(* IEC 61131-3 sources: structured-text/samples/unsupported/arrays, 10 files *)

(* ---- f.4.st ---- *)
FUNCTION_BLOCK STACK_INT
  VAR_INPUT PUSH, POP: BOOL;
            R1 : BOOL ;
            IN : INT ;
            N  : INT ;
  END_VAR
  VAR_OUTPUT EMPTY : BOOL := 1 ;
             OFLO  : BOOL := 0 ;
             OUT   : INT  := 0 ;
  END_VAR
  VAR STK : ARRAY[0..127] OF INT;
      NI : INT :=128  ;
      PTR : INT := -1 ;
  END_VAR

    IF R1 THEN
       OFLO := 0; EMPTY := 1; PTR := -1;
       NI := LIMIT (MN:=1,IN:=N,MX:=128); OUT := 0;
    ELSIF POP & NOT EMPTY THEN
       OFLO := 0; PTR := PTR-1; EMPTY := PTR < 0;
       IF EMPTY THEN OUT := 0;
       ELSE OUT := STK[PTR];
       END_IF ;
    ELSIF PUSH & NOT OFLO THEN
       EMPTY := 0; PTR := PTR+1; OFLO := (PTR = NI);
       IF NOT OFLO THEN OUT := IN ; STK[PTR] := IN;
       ELSE OUT := 0;
       END_IF ;
    END_IF ;
END_FUNCTION_BLOCK

(* ---- f.6.11.st ---- *)
FUNCTION_BLOCK DIFFEQ
   VAR_INPUT
     RUN : BOOL ;
     XIN : REAL ;
     A : ARRAY[1..127] OF REAL ;
     M : INT ;
     B : ARRAY[0..127] OF REAL ;
     N : INT ;
   END_VAR
   VAR_OUTPUT XOUT : REAL := 0.0 ; END_VAR
   VAR
     XI : ARRAY [0..127] OF REAL ;
     XO : ARRAY [0..127] OF REAL ;
     I : INT ;
   END_VAR
   XO[0] := XOUT ; XI[0] := XIN ;
   XOUT := B[0] * XIN ;
   IF RUN THEN
      FOR I := M TO 1 BY -1 DO
          XOUT := XOUT + A[I] * XO[I] ; XO[I] := XO[I-1];
      END_FOR;
      FOR I := N TO 1 BY -1 DO
          XOUT := XOUT + B[I] * XI[I] ; XI[I] := XI[I-1];
      END_FOR;
   ELSE
      FOR I := 1 TO M DO XO[I] := 0.0; END_FOR;
      FOR I := 1 TO N DO XI[I] := 0.0; END_FOR;
   END_IF ;
 END_FUNCTION_BLOCK

(* ---- f.6.2.st ---- *)
FUNCTION_BLOCK DELAY
  VAR_INPUT
    RUN : BOOL ;
    XIN : REAL ;
    N   : INT ;
  END_VAR
  VAR_OUTPUT XOUT : REAL; END_VAR
  VAR X : ARRAY [0..127]
               OF REAL;
      I, IXIN, IXOUT : INT := 0;
  END_VAR
  IF RUN THEN IXIN := MOD(IXIN + 1, 128) ; X[IXIN] := XIN ;
              IXOUT := MOD(IXOUT + 1, 128) ; XOUT := X[IXOUT];
  ELSE XOUT := XIN ; IXIN := N ; IXOUT := 0;
       FOR I := 0 TO N DO X[I] := XIN; END_FOR;
  END_IF ;
END_FUNCTION_BLOCK

(* ---- t17-4.st ---- *)
PROGRAM Test
	VAR
		INARY AT %IW6 ;
 		ARRAY [0..9] OF INT;
	END_VAR
END_PROGRAM

(* ---- t17-6.st ---- *)
PROGRAM Test
	VAR THREE :
		ARRAY[1..5,1..10,1..8] OF INT;
	END_VAR
END_PROGRAM

(* ---- t17-7.st ---- *)
PROGRAM Test
	VAR RETAIN RTBT:
  		ARRAY[1..2,1..3] OF INT;
	END_VAR
END_PROGRAM

(* ---- t18-4.st ---- *)
PROGRAM Test
	VAR OUTARY AT %QW6 :
 		ARRAY[0..9] OF INT := [10(1)];
	END_VAR
END_PROGRAM

(* ---- t18-6.st ---- *)
PROGRAM Test
	VAR
		BITS : ARRAY[0..7]
			OF BOOL := [1,1,0,0,0,1,0,0] ;
	  	TBT : ARRAY [1..2,1..3]
	        OF INT := [1,2,3(4),6] ;
	END_VAR
END_PROGRAM

(* ---- t18-7.st ---- *)
PROGRAM Test
	VAR RETAIN RTBT :
  		ARRAY(1..2,1..3) OF INT
      		:= [1,2,3(4)];
	END_VAR
END_PROGRAM

(* ---- t18-8.st ---- *)
PROGRAM Test
	VAR MODULE_8_CONFIG:
	  ANALOG_16_INPUT_CONFIGURATION :=
	    (SIGNAL_TYPE := DIFFERENTIAL,
	      CHANNEL
	        := [4((RANGE := UNIPOLAR_1_5V)),
	            (RANGE:= BIPOLAR_10_V,
	             MIN_SCALE := 0,
	             MAX_SCALE := 500)]);
	END_VAR
END_PROGRAM
